// Characterisation tests of HalfBROT.FB_HydraulicsControl (HalfBROT#32 step 3) through the I/O structs and the command methods
// (#30, #31): start-up, the brake (pressure delay, clearing, pressure loss, CloseBrake, pump stop, azimuth limit), the manual
// brake re-arm of #31, and the latched errors that need no more than 13 s. They pin what the block does today, they are
// not a specification. Every test owns a rig (FB_HydraulicsRig, a plant behind the structs) and runs over many PLC cycles;
// the block timers run on the system time, so the tests take real time (the longest about 15 s). The suction and
// pressure watchdogs are shortened through tSuctionWatchdog and tPressureWatchdog.
FUNCTION_BLOCK FB_HydraulicsControl_Tests EXTENDS FB_TestBase
VAR
END_VAR

Idle_Everything_Off();
Enable_Runs_Pump();
Open_Brake_After_Pressure_Delay();
No_Clearing_Keeps_Brake_Closed();
Pressure_Loss_Closes_Brake_Auto_Reopens();
CloseBrake_Closes_And_Ends_Request();
Pump_Stop_Closes_Brake();
Azimuth_Limit_Closes_Brake();
Manual_Brake_Stays_Closed_After_Pressure_Loss();
Manual_Brake_Reopens_After_Switch_Off_On();
Manual_Switch_Off_Closes_Brake();
Manual_Brake_Stays_Closed_After_Pump_Restart();
Oil_Low_Is_Error_Until_Reset();
Hydraulics_Watchdog_Is_Error();
Suction_Without_Feedback_Is_Error();
Missing_Pressure_Is_Error();
Main_Pump_Without_Feedback_Is_Error();

// No request, healthy sensors: no pump, no brake, no error, no starter reset.
METHOD PRIVATE Idle_Everything_Off
VAR_INST
	rig		: FB_HydraulicsRig;
	nStep	: INT;
	bViol	: BOOL;
END_VAR
TEST('Idle_Everything_Off');
sCurrent := 'Idle_Everything_Off: ';
IF nStep >= 90 THEN
	RETURN;
END_IF
rig.Scan();
IF rig.nScans >= 5 THEN
	Check(NOT rig.stOut.bOilPumpEnable, 'no pump enable');
	Check(NOT rig.stOut.bOilSuctionEnable, 'no suction enable');
	Check(NOT rig.stOut.bBrakeAzEl, 'brake output off');
	Check(NOT rig.fb.bError, 'no error with healthy sensors');
	Check(rig.fb.PumpState = HalfBROT.E_PumpState.Off, 'pump state Off');
	Check(rig.fb.bBrakeClosed AND NOT rig.fb.bBrakeOpen, 'brake reported closed');
	Check(rig.fb.BrakeState = HalfBROT.E_BrakeState.Closed, 'brake state Closed');
	Check(NOT rig.stOut.bResetOilPump AND NOT rig.stOut.bResetSuctionPump, 'no starter reset');
		nStep := 99;
		TEST_FINISHED();
END_IF
END_METHOD

// Enable starts the pump; the plant reports it running with pressure; the brake is not opened by the pump start.
METHOD PRIVATE Enable_Runs_Pump
VAR_INST
	rig		: FB_HydraulicsRig;
	nStep	: INT;
	bViol	: BOOL;
END_VAR
TEST('Enable_Runs_Pump');
sCurrent := 'Enable_Runs_Pump: ';
IF nStep >= 90 THEN
	RETURN;
END_IF
rig.Scan();
CASE nStep OF
0:
	rig.SetEnable(TRUE);
	rig.StepStart();
	nStep := 10;
10:
	IF rig.nStepScans >= 6 THEN
		Check(rig.fb.Enable, 'Enable reads back');
		Check(rig.stOut.bOilPumpEnable, 'pump enable output');
		Check(rig.fb.PumpRunning AND rig.fb.OilPressureOK, 'pump running and pressure reported');
		Check(rig.fb.PumpState = HalfBROT.E_PumpState.Running, 'pump state Running');
		Check(NOT rig.fb.Error, 'no error');
		Check(NOT rig.stOut.bBrakeAzEl, 'the pump start does not open the brake');
		nStep := 99;
		TEST_FINISHED();
	END_IF
END_CASE
END_METHOD

// OpenBrake() each scan: the brake output comes about 3 s after the pressure, the report 1 s after the output.
METHOD PRIVATE Open_Brake_After_Pressure_Delay
VAR_INST
	rig		: FB_HydraulicsRig;
	nStep	: INT;
	bViol	: BOOL;
END_VAR
TEST('Open_Brake_After_Pressure_Delay');
sCurrent := 'Open_Brake_After_Pressure_Delay: ';
IF nStep >= 90 THEN
	RETURN;
END_IF
rig.Scan();
CASE nStep OF
0:
	rig.bClearing := TRUE;
	rig.bAuto := TRUE;
	rig.SetEnable(TRUE);
	rig.StepStart();
	nStep := 10;
10:
	IF rig.StepTime(T#1S) THEN
		Check(NOT rig.stOut.bBrakeAzEl, 'no brake output during the pressure delay');
		nStep := 20;
	END_IF
20:
	IF rig.stOut.bBrakeAzEl THEN
		Check(rig.StepTime(T#2S500MS) AND NOT rig.StepTime(T#4S), 'the brake output comes about 3 s after the start');
		Check(NOT rig.fb.bBrakeOpen, 'open is reported 1 s after the output, not with it');
		Check(rig.fb.BrakeState = HalfBROT.E_BrakeState.Opening, 'brake state Opening while the output is on and not reported');
		rig.StepStart();
		nStep := 30;
	ELSIF rig.StepTime(T#6S) THEN
		Check(FALSE, 'the brake output never came');
		nStep := 99;
		TEST_FINISHED();
	END_IF
30:
	IF rig.fb.bBrakeOpen THEN
		Check(rig.StepTime(T#800MS) AND NOT rig.StepTime(T#2S), 'open is reported about 1 s after the output');
		Check(rig.fb.BrakeOpen AND NOT rig.fb.bBrakeClosed, 'BrakeOpen property and bBrakeClosed agree');
		Check(rig.fb.BrakeState = HalfBROT.E_BrakeState.Open, 'brake state Open when reported');
		nStep := 99;
		TEST_FINISHED();
	ELSIF rig.StepTime(T#3S) THEN
		Check(FALSE, 'open was never reported');
		nStep := 99;
		TEST_FINISHED();
	END_IF
END_CASE
END_METHOD

// Without bBrakeClearing the brake is not opened although it is requested and the pressure is there.
METHOD PRIVATE No_Clearing_Keeps_Brake_Closed
VAR_INST
	rig		: FB_HydraulicsRig;
	nStep	: INT;
	bViol	: BOOL;
END_VAR
TEST('No_Clearing_Keeps_Brake_Closed');
sCurrent := 'No_Clearing_Keeps_Brake_Closed: ';
IF nStep >= 90 THEN
	RETURN;
END_IF
rig.Scan();
CASE nStep OF
0:
	rig.bClearing := FALSE;
	rig.bAuto := TRUE;
	rig.SetEnable(TRUE);
	rig.StepStart();
	nStep := 10;
10:
	bViol := bViol OR rig.stOut.bBrakeAzEl OR rig.fb.bBrakeOpen;
	IF rig.StepTime(T#4S) THEN
		Check(NOT bViol, 'the brake stays closed without the clearing');
		Check(rig.fb.PumpRunning AND rig.fb.OilPressureOK, 'pump running with pressure');
		nStep := 99;
		TEST_FINISHED();
	END_IF
END_CASE
END_METHOD

// Pressure loss closes the brake after the 2 s debounce; with the automatic request still there it opens again after the pressure delay.
METHOD PRIVATE Pressure_Loss_Closes_Brake_Auto_Reopens
VAR_INST
	rig		: FB_HydraulicsRig;
	nStep	: INT;
	bViol	: BOOL;
END_VAR
TEST('Pressure_Loss_Closes_Brake_Auto_Reopens');
sCurrent := 'Pressure_Loss_Closes_Brake_Auto_Reopens: ';
IF nStep >= 90 THEN
	RETURN;
END_IF
rig.Scan();
CASE nStep OF
0:
	rig.bClearing := TRUE;
	rig.bAuto := TRUE;
	rig.SetEnable(TRUE);
	rig.StepStart();
	nStep := 10;
10:
	IF rig.fb.bBrakeOpen THEN
		rig.bPressure := FALSE;
		rig.StepStart();
		nStep := 20;
	ELSIF rig.StepTime(T#8S) THEN
		Check(FALSE, 'the brake never opened');
		nStep := 99;
		TEST_FINISHED();
	END_IF
20:
	IF NOT rig.stOut.bBrakeAzEl THEN
		Check(rig.StepTime(T#1S500MS), 'the brake holds during the 2 s debounce');
		Check(NOT rig.fb.bBrakeOpen, 'closed is reported');
		Check(rig.stOut.bOilPumpEnable, 'the pump enable stays');
		rig.bPressure := TRUE;
		rig.StepStart();
		nStep := 30;
	ELSIF rig.StepTime(T#4S) THEN
		Check(FALSE, 'the brake did not close on the pressure loss');
		nStep := 99;
		TEST_FINISHED();
	END_IF
30:
	IF rig.stOut.bBrakeAzEl THEN
		Check(rig.StepTime(T#2S), 'the brake opens again only after the pressure delay');
		nStep := 99;
		TEST_FINISHED();
	ELSIF rig.StepTime(T#6S) THEN
		Check(FALSE, 'the automatic request did not open the brake again');
		nStep := 99;
		TEST_FINISHED();
	END_IF
END_CASE
END_METHOD

// CloseBrake() closes the brake at once and the request ends: no automatic re-open without OpenBrake().
METHOD PRIVATE CloseBrake_Closes_And_Ends_Request
VAR_INST
	rig		: FB_HydraulicsRig;
	nStep	: INT;
	bViol	: BOOL;
END_VAR
TEST('CloseBrake_Closes_And_Ends_Request');
sCurrent := 'CloseBrake_Closes_And_Ends_Request: ';
IF nStep >= 90 THEN
	RETURN;
END_IF
rig.Scan();
CASE nStep OF
0:
	rig.bClearing := TRUE;
	rig.bAuto := TRUE;
	rig.SetEnable(TRUE);
	rig.StepStart();
	nStep := 10;
10:
	IF rig.fb.bBrakeOpen THEN
		rig.bAuto := FALSE;
		rig.fb.CloseBrake();
		rig.StepStart();
		nStep := 20;
	ELSIF rig.StepTime(T#8S) THEN
		Check(FALSE, 'the brake never opened');
		nStep := 99;
		TEST_FINISHED();
	END_IF
20:
	IF NOT rig.stOut.bBrakeAzEl THEN
		Check(NOT rig.StepTime(T#300MS), 'the brake output drops at once');
		Check(NOT rig.fb.bBrakeOpen, 'closed is reported');
		Check(rig.fb.BrakeState = HalfBROT.E_BrakeState.Closed, 'brake state Closed after the close');
		rig.StepStart();
		nStep := 30;
	ELSIF rig.StepTime(T#1S) THEN
		Check(FALSE, 'CloseBrake() did not close the brake');
		nStep := 99;
		TEST_FINISHED();
	END_IF
30:
	bViol := bViol OR rig.stOut.bBrakeAzEl;
	IF rig.StepTime(T#4S) THEN
		Check(NOT bViol, 'the brake stays closed with the pressure there');
		nStep := 99;
		TEST_FINISHED();
	END_IF
END_CASE
END_METHOD

// ManualStopPump drops the pump enable; with the pump the brake closes.
METHOD PRIVATE Pump_Stop_Closes_Brake
VAR_INST
	rig		: FB_HydraulicsRig;
	nStep	: INT;
	bViol	: BOOL;
END_VAR
TEST('Pump_Stop_Closes_Brake');
sCurrent := 'Pump_Stop_Closes_Brake: ';
IF nStep >= 90 THEN
	RETURN;
END_IF
rig.Scan();
CASE nStep OF
0:
	rig.bClearing := TRUE;
	rig.bAuto := TRUE;
	rig.SetEnable(TRUE);
	rig.StepStart();
	nStep := 10;
10:
	IF rig.fb.bBrakeOpen THEN
		rig.bAuto := FALSE;
		rig.SetStopPump(TRUE);
		rig.StepStart();
		nStep := 20;
	ELSIF rig.StepTime(T#8S) THEN
		Check(FALSE, 'the brake never opened');
		nStep := 99;
		TEST_FINISHED();
	END_IF
20:
	IF NOT rig.stOut.bBrakeAzEl THEN
		Check(NOT rig.StepTime(T#300MS), 'the brake output drops with the pump');
		Check(NOT rig.stOut.bOilPumpEnable, 'pump enable off');
		Check(NOT rig.fb.bBrakeOpen, 'closed is reported');
		nStep := 99;
		TEST_FINISHED();
	ELSIF rig.StepTime(T#1S) THEN
		Check(FALSE, 'the pump stop did not close the brake');
		nStep := 99;
		TEST_FINISHED();
	END_IF
END_CASE
END_METHOD

// The azimuth limit switch closes the brake and holds it closed while it is active, although the request goes on.
METHOD PRIVATE Azimuth_Limit_Closes_Brake
VAR_INST
	rig		: FB_HydraulicsRig;
	nStep	: INT;
	bViol	: BOOL;
END_VAR
TEST('Azimuth_Limit_Closes_Brake');
sCurrent := 'Azimuth_Limit_Closes_Brake: ';
IF nStep >= 90 THEN
	RETURN;
END_IF
rig.Scan();
CASE nStep OF
0:
	rig.bClearing := TRUE;
	rig.bAuto := TRUE;
	rig.SetEnable(TRUE);
	rig.StepStart();
	nStep := 10;
10:
	IF rig.fb.bBrakeOpen THEN
		rig.bAzLimit := TRUE;
		rig.StepStart();
		nStep := 20;
	ELSIF rig.StepTime(T#8S) THEN
		Check(FALSE, 'the brake never opened');
		nStep := 99;
		TEST_FINISHED();
	END_IF
20:
	IF NOT rig.stOut.bBrakeAzEl THEN
		Check(NOT rig.StepTime(T#300MS), 'the brake output drops at once');
		rig.StepStart();
		nStep := 30;
	ELSIF rig.StepTime(T#1S) THEN
		Check(FALSE, 'the azimuth limit did not close the brake');
		nStep := 99;
		TEST_FINISHED();
	END_IF
30:
	bViol := bViol OR rig.stOut.bBrakeAzEl;
	IF rig.StepTime(T#4S) THEN
		Check(NOT bViol, 'the brake stays closed while the limit is active');
		nStep := 99;
		TEST_FINISHED();
	END_IF
END_CASE
END_METHOD

// #31: the cabinet switch opens the brake once; after a pressure loss it stays closed while the switch stays on, with the pressure back.
METHOD PRIVATE Manual_Brake_Stays_Closed_After_Pressure_Loss
VAR_INST
	rig		: FB_HydraulicsRig;
	nStep	: INT;
	bViol	: BOOL;
END_VAR
TEST('Manual_Brake_Stays_Closed_After_Pressure_Loss');
sCurrent := 'Manual_Brake_Stays_Closed_After_Pressure_Loss: ';
IF nStep >= 90 THEN
	RETURN;
END_IF
rig.Scan();
CASE nStep OF
0:
	// the pump runs first: a switch edge before the pump runs is dropped by the block (the request is cleared while the pump is off)
	rig.bManual := TRUE;
	rig.SetEnable(TRUE);
	rig.StepStart();
	nStep := 5;
5:
	IF rig.StepTime(T#500MS) THEN
		rig.bSwitch := TRUE;
		rig.StepStart();
		nStep := 10;
	END_IF
10:
	IF rig.fb.bBrakeOpen THEN
		Check(rig.stOut.bBrakeAzEl, 'the switch opened the brake');
		rig.bPressure := FALSE;
		rig.StepStart();
		nStep := 20;
	ELSIF rig.StepTime(T#8S) THEN
		Check(FALSE, 'the brake never opened');
		nStep := 99;
		TEST_FINISHED();
	END_IF
20:
	IF NOT rig.stOut.bBrakeAzEl THEN
		Check(rig.StepTime(T#1S500MS), 'the brake holds during the 2 s debounce');
		rig.bPressure := TRUE;
		bViol := FALSE;
		rig.StepStart();
		nStep := 30;
	ELSIF rig.StepTime(T#4S) THEN
		Check(FALSE, 'the brake did not close on the pressure loss');
		nStep := 99;
		TEST_FINISHED();
	END_IF
30:
	bViol := bViol OR rig.stOut.bBrakeAzEl;
	IF rig.StepTime(T#4S500MS) THEN
		Check(rig.fb.bOilPressureOK AND rig.fb.PumpRunning, 'pressure is back');
		Check(NOT bViol, 'the brake is not opened again while the switch stays on');
		nStep := 99;
		TEST_FINISHED();
	END_IF
END_CASE
END_METHOD

// #31: after CloseBrake() the brake stays closed while the switch stays on; switch off and on opens it again.
METHOD PRIVATE Manual_Brake_Reopens_After_Switch_Off_On
VAR_INST
	rig		: FB_HydraulicsRig;
	nStep	: INT;
	bViol	: BOOL;
END_VAR
TEST('Manual_Brake_Reopens_After_Switch_Off_On');
sCurrent := 'Manual_Brake_Reopens_After_Switch_Off_On: ';
IF nStep >= 90 THEN
	RETURN;
END_IF
rig.Scan();
CASE nStep OF
0:
	// the pump runs first: a switch edge before the pump runs is dropped by the block (the request is cleared while the pump is off)
	rig.bManual := TRUE;
	rig.SetEnable(TRUE);
	rig.StepStart();
	nStep := 5;
5:
	IF rig.StepTime(T#500MS) THEN
		rig.bSwitch := TRUE;
		rig.StepStart();
		nStep := 10;
	END_IF
10:
	IF rig.fb.bBrakeOpen THEN
		rig.fb.CloseBrake();
		rig.StepStart();
		nStep := 20;
	ELSIF rig.StepTime(T#8S) THEN
		Check(FALSE, 'the brake never opened');
		nStep := 99;
		TEST_FINISHED();
	END_IF
20:
	IF NOT rig.stOut.bBrakeAzEl THEN
		Check(NOT rig.StepTime(T#300MS), 'CloseBrake() closes at once');
		bViol := FALSE;
		rig.StepStart();
		nStep := 30;
	ELSIF rig.StepTime(T#1S) THEN
		Check(FALSE, 'CloseBrake() did not close the brake');
		nStep := 99;
		TEST_FINISHED();
	END_IF
30:
	bViol := bViol OR rig.stOut.bBrakeAzEl;
	IF rig.StepTime(T#4S) THEN
		Check(NOT bViol, 'the brake stays closed while the switch stays on');
		rig.bSwitch := FALSE;
		rig.StepStart();
		nStep := 40;
	END_IF
40:
	IF rig.StepTime(T#500MS) THEN
		Check(NOT rig.stOut.bBrakeAzEl, 'the brake is closed with the switch off');
		rig.bSwitch := TRUE;
		rig.StepStart();
		nStep := 50;
	END_IF
50:
	IF rig.stOut.bBrakeAzEl THEN
		Check(NOT rig.StepTime(T#1S), 'the switch off and on opens the brake at once, the pressure delay has long run out');
		nStep := 99;
		TEST_FINISHED();
	ELSIF rig.StepTime(T#6S) THEN
		Check(FALSE, 'the brake did not open again after the switch went off and on');
		nStep := 99;
		TEST_FINISHED();
	END_IF
END_CASE
END_METHOD

// The permission: switch off closes the brake at once (bBrakeClearing) and ends the request.
METHOD PRIVATE Manual_Switch_Off_Closes_Brake
VAR_INST
	rig		: FB_HydraulicsRig;
	nStep	: INT;
	bViol	: BOOL;
END_VAR
TEST('Manual_Switch_Off_Closes_Brake');
sCurrent := 'Manual_Switch_Off_Closes_Brake: ';
IF nStep >= 90 THEN
	RETURN;
END_IF
rig.Scan();
CASE nStep OF
0:
	// the pump runs first: a switch edge before the pump runs is dropped by the block (the request is cleared while the pump is off)
	rig.bManual := TRUE;
	rig.SetEnable(TRUE);
	rig.StepStart();
	nStep := 5;
5:
	IF rig.StepTime(T#500MS) THEN
		rig.bSwitch := TRUE;
		rig.StepStart();
		nStep := 10;
	END_IF
10:
	IF rig.fb.bBrakeOpen THEN
		rig.bSwitch := FALSE;
		rig.StepStart();
		nStep := 20;
	ELSIF rig.StepTime(T#8S) THEN
		Check(FALSE, 'the brake never opened');
		nStep := 99;
		TEST_FINISHED();
	END_IF
20:
	IF NOT rig.stOut.bBrakeAzEl THEN
		Check(NOT rig.StepTime(T#300MS), 'the brake output drops at once');
		Check(NOT rig.fb.bBrakeOpen, 'closed is reported');
		Check(rig.fb.BrakeState = HalfBROT.E_BrakeState.Closed, 'brake state Closed after the close');
		nStep := 99;
		TEST_FINISHED();
	ELSIF rig.StepTime(T#1S) THEN
		Check(FALSE, 'the switch off did not close the brake');
		nStep := 99;
		TEST_FINISHED();
	END_IF
END_CASE
END_METHOD

// #31: a pump stop closes the brake; the pump runs again with the switch still on: the brake stays closed.
METHOD PRIVATE Manual_Brake_Stays_Closed_After_Pump_Restart
VAR_INST
	rig		: FB_HydraulicsRig;
	nStep	: INT;
	bViol	: BOOL;
END_VAR
TEST('Manual_Brake_Stays_Closed_After_Pump_Restart');
sCurrent := 'Manual_Brake_Stays_Closed_After_Pump_Restart: ';
IF nStep >= 90 THEN
	RETURN;
END_IF
rig.Scan();
CASE nStep OF
0:
	// the pump runs first: a switch edge before the pump runs is dropped by the block (the request is cleared while the pump is off)
	rig.bManual := TRUE;
	rig.SetEnable(TRUE);
	rig.StepStart();
	nStep := 5;
5:
	IF rig.StepTime(T#500MS) THEN
		rig.bSwitch := TRUE;
		rig.StepStart();
		nStep := 10;
	END_IF
10:
	IF rig.fb.bBrakeOpen THEN
		rig.SetStopPump(TRUE);
		rig.StepStart();
		nStep := 20;
	ELSIF rig.StepTime(T#8S) THEN
		Check(FALSE, 'the brake never opened');
		nStep := 99;
		TEST_FINISHED();
	END_IF
20:
	IF NOT rig.stOut.bBrakeAzEl THEN
		Check(NOT rig.StepTime(T#300MS), 'the pump stop closes the brake at once');
		rig.StepStart();
		nStep := 30;
	ELSIF rig.StepTime(T#1S) THEN
		Check(FALSE, 'the pump stop did not close the brake');
		nStep := 99;
		TEST_FINISHED();
	END_IF
30:
	IF rig.StepTime(T#500MS) THEN
		rig.SetStopPump(FALSE);
		bViol := FALSE;
		rig.StepStart();
		nStep := 40;
	END_IF
40:
	bViol := bViol OR rig.stOut.bBrakeAzEl;
	IF rig.StepTime(T#4S500MS) THEN
		Check(rig.fb.PumpRunning AND rig.fb.OilPressureOK, 'the pump runs again with pressure');
		Check(NOT bViol, 'the brake is not opened again while the switch stays on');
		nStep := 99;
		TEST_FINISHED();
	END_IF
END_CASE
END_METHOD

// Oil low is a latched error that stops the pump; Reset() clears it once the oil is back and the pump starts again (Enable is still set).
METHOD PRIVATE Oil_Low_Is_Error_Until_Reset
VAR_INST
	rig		: FB_HydraulicsRig;
	nStep	: INT;
	bViol	: BOOL;
END_VAR
TEST('Oil_Low_Is_Error_Until_Reset');
sCurrent := 'Oil_Low_Is_Error_Until_Reset: ';
IF nStep >= 90 THEN
	RETURN;
END_IF
rig.Scan();
CASE nStep OF
0:
	rig.SetEnable(TRUE);
	rig.StepStart();
	nStep := 10;
10:
	IF rig.nStepScans >= 5 THEN
		rig.stIn.bOilLow := FALSE;
		rig.StepStart();
		nStep := 20;
	END_IF
20:
	IF rig.nStepScans >= 3 THEN
		Check(rig.fb.Error AND rig.fb.bOilLow, 'oil low is an error');
		Check(rig.fb.PumpState = HalfBROT.E_PumpState.Error, 'pump state Error');
		Check(NOT rig.stOut.bOilPumpEnable, 'the error stops the pump');
		rig.stIn.bOilLow := TRUE;
		rig.StepStart();
		nStep := 30;
	END_IF
30:
	IF rig.nStepScans >= 3 THEN
		Check(rig.fb.Error, 'the error stays latched with the oil back');
		rig.fb.Reset();
		rig.StepStart();
		nStep := 40;
	END_IF
40:
	IF rig.nStepScans >= 4 THEN
		Check(NOT rig.fb.Error, 'Reset() clears the error');
		Check(rig.stOut.bOilPumpEnable, 'the pump starts again, Enable is still set');
		Check(rig.fb.PumpState = HalfBROT.E_PumpState.Running, 'pump state Running again after Reset()');
		nStep := 99;
		TEST_FINISHED();
	END_IF
END_CASE
END_METHOD

// The pump running without the suction pump for tHydraulicsWatchdog (1 s here, 140 s default, #10) is a latched error.
METHOD PRIVATE Hydraulics_Watchdog_Is_Error
VAR_INST
	rig		: FB_HydraulicsRig;
	nStep	: INT;
	bViol	: BOOL;
END_VAR
TEST('Hydraulics_Watchdog_Is_Error');
sCurrent := 'Hydraulics_Watchdog_Is_Error: ';
IF nStep >= 90 THEN
	RETURN;
END_IF
rig.Scan();
CASE nStep OF
0:
	rig.tHydraulicsWatchdog := T#1S;
	rig.bSuctionFollows := FALSE;
	rig.SetEnable(TRUE);
	rig.StepStart();
	nStep := 10;
10:
	bViol := bViol OR rig.fb.bHydraulicsFailure;
	IF rig.fb.Error THEN
		Check(rig.StepTime(T#800MS), 'not before the configured time');
		Check(bViol, 'the hydraulics failure was reported');
		Check(NOT rig.stOut.bOilPumpEnable, 'the error stops the pump');
		nStep := 99;
		TEST_FINISHED();
	ELSIF rig.StepTime(T#4S) THEN
		Check(FALSE, 'no hydraulics failure');
		nStep := 99;
		TEST_FINISHED();
	END_IF
END_CASE
END_METHOD

// The suction enable (manual start) without the run feedback for tSuctionWatchdog (1 s here, 15 s default) is a latched error.
METHOD PRIVATE Suction_Without_Feedback_Is_Error
VAR_INST
	rig		: FB_HydraulicsRig;
	nStep	: INT;
	bViol	: BOOL;
END_VAR
TEST('Suction_Without_Feedback_Is_Error');
sCurrent := 'Suction_Without_Feedback_Is_Error: ';
IF nStep >= 90 THEN
	RETURN;
END_IF
rig.Scan();
CASE nStep OF
0:
	rig.tSuctionWatchdog := T#1S;
	rig.bSuctionFollows := FALSE;
	rig.SetSuction(TRUE);
	rig.StepStart();
	nStep := 10;
10:
	bViol := bViol OR rig.fb.bSuctionFailure;
	IF rig.fb.Error THEN
		Check(rig.stOut.bOilSuctionEnable, 'the suction enable was on');
		Check(rig.StepTime(T#800MS), 'not before the configured time');
		Check(bViol, 'the suction failure was reported');
		nStep := 99;
		TEST_FINISHED();
	ELSIF rig.StepTime(T#4S) THEN
		Check(FALSE, 'no suction failure');
		nStep := 99;
		TEST_FINISHED();
	END_IF
END_CASE
END_METHOD

// The pump enabled without oil pressure for tPressureWatchdog (1 s here, 30 s default) is a latched error that stops the pump.
METHOD PRIVATE Missing_Pressure_Is_Error
VAR_INST
	rig		: FB_HydraulicsRig;
	nStep	: INT;
	bViol	: BOOL;
END_VAR
TEST('Missing_Pressure_Is_Error');
sCurrent := 'Missing_Pressure_Is_Error: ';
IF nStep >= 90 THEN
	RETURN;
END_IF
rig.Scan();
CASE nStep OF
0:
	rig.tPressureWatchdog := T#1S;
	rig.bPressure := FALSE;
	rig.SetEnable(TRUE);
	rig.StepStart();
	nStep := 10;
10:
	bViol := bViol OR rig.fb.bPressureFailure;
	IF rig.fb.Error THEN
		Check(rig.StepTime(T#800MS), 'not before the configured time');
		Check(bViol, 'the pressure failure was reported');
		Check(NOT rig.stOut.bOilPumpEnable, 'the error stops the pump');
		nStep := 99;
		TEST_FINISHED();
	ELSIF rig.StepTime(T#4S) THEN
		Check(FALSE, 'no pressure failure');
		nStep := 99;
		TEST_FINISHED();
	END_IF
END_CASE
END_METHOD

// No run feedback 10 s after the pump enable is a latched error (main pump failure).
METHOD PRIVATE Main_Pump_Without_Feedback_Is_Error
VAR_INST
	rig		: FB_HydraulicsRig;
	nStep	: INT;
	bViol	: BOOL;
END_VAR
TEST('Main_Pump_Without_Feedback_Is_Error');
sCurrent := 'Main_Pump_Without_Feedback_Is_Error: ';
IF nStep >= 90 THEN
	RETURN;
END_IF
rig.Scan();
CASE nStep OF
0:
	rig.bPumpFollows := FALSE;
	rig.SetEnable(TRUE);
	rig.StepStart();
	nStep := 10;
10:
	bViol := bViol OR rig.fb.bMainPumpFailure;
	IF rig.fb.Error THEN
		Check(rig.StepTime(T#9S500MS), 'not before the 10 s');
		Check(bViol, 'the main pump failure was reported');
		Check(NOT rig.stOut.bOilPumpEnable, 'the error stops the pump');
		nStep := 99;
		TEST_FINISHED();
	ELSIF rig.StepTime(T#13S) THEN
		Check(FALSE, 'no main pump failure');
		nStep := 99;
		TEST_FINISHED();
	END_IF
END_CASE
END_METHOD

END_FUNCTION_BLOCK

(* stored: Version 1.1.0.1, ProductVersion 3.1.4024.15
   POU FB_HydraulicsControl_Tests: Id {d102baa1-bfde-5915-adf5-4a2f2c8fb59d}, SpecialFunc None
   Method Idle_Everything_Off: Id {ae63437a-f211-52ef-a794-791e9d874db8}
   Method Enable_Runs_Pump: Id {c3347adc-7271-5702-9f14-c4d806e5384d}
   Method Open_Brake_After_Pressure_Delay: Id {4823ab7a-7d97-5ca4-879f-8dd315ac05a4}
   Method No_Clearing_Keeps_Brake_Closed: Id {65246b8a-191b-56f8-87c9-56a638e8452d}
   Method Pressure_Loss_Closes_Brake_Auto_Reopens: Id {ceb24780-919e-518e-b9b6-7a73071a85e8}
   Method CloseBrake_Closes_And_Ends_Request: Id {d05ec3f7-f71e-5ad3-8ac8-675addc014a6}
   Method Pump_Stop_Closes_Brake: Id {b2541adb-c4f8-5bc5-bdbd-2133fdafcbf7}
   Method Azimuth_Limit_Closes_Brake: Id {1042741a-a56a-553b-99e2-8f1ddb3a23a2}
   Method Manual_Brake_Stays_Closed_After_Pressure_Loss: Id {69151a09-53e3-5aba-8f12-4e584c9ffdf8}
   Method Manual_Brake_Reopens_After_Switch_Off_On: Id {1e3f6eef-f200-589f-a4c3-9b09506881cd}
   Method Manual_Switch_Off_Closes_Brake: Id {ec6a1f02-9aa3-5941-a3a9-899a208b86fa}
   Method Manual_Brake_Stays_Closed_After_Pump_Restart: Id {de6329f8-21ed-55dc-b182-00ec3d3e3509}
   Method Oil_Low_Is_Error_Until_Reset: Id {50b3c179-5e93-5f1e-9dab-809e9ea04152}
   Method Hydraulics_Watchdog_Is_Error: Id {dc55646e-87ae-5b84-a5bd-27ab2874fd35}
   Method Suction_Without_Feedback_Is_Error: Id {40af0bb4-28fd-5a42-ab7e-694edfb5dd03}
   Method Missing_Pressure_Is_Error: Id {6b86aa9c-2d68-589f-94f5-02d5eeeffca0}
   Method Main_Pump_Without_Feedback_Is_Error: Id {44ac1229-1e49-55b7-81df-aa7992b702da} *)
